// TIA Portal V20 export
// export: Created 2026-10-11T05:25:30.6576364Z, ExportSetting WithDefaults, DisplayName Totally Integrated Automation Portal, DisplayVersion V20, DisplayName TIA Portal Openness, DisplayVersion V20, DisplayName TIA Portal Teamcenter Gateway, DisplayVersion V20, DisplayName TIA Portal Version Control Interface, DisplayVersion V20, DisplayName SINAMICS Startdrive Advanced, DisplayVersion V20 SP1 Update 2, DisplayName SINAMICS Startdrive G110M, G120, G120C, G120D, G120P, G115D, DisplayVersion V20 SP1 Update 2, DisplayName SINAMICS Startdrive G130, G150, S120, S150, SINAMICS MV, G220, S200, S210, DisplayVersion V20 SP1 Update 2, DisplayName STEP 7 Professional, DisplayVersion V20, DisplayName STEP 7 Safety, DisplayVersion V20, DisplayName WinCC Basic/Comfort/Advanced, DisplayVersion V20, DisplayName WinCC Professional, DisplayVersion V20, DisplayName WinCC Unified, DisplayVersion V20
FUNCTION "FRK_PartReceived" : Bool   // FC38, SCL
{ S7_Optimized_Access := 'TRUE' }
VERSION : 0.1
// stored: AutoNumber true, IsIECCheckEnabled false, SetENOAutomatically false, UDAEnableTagReadback false
   VAR_IN_OUT
      Core : "FRK_Core";
      Unit : "FRK_Unit";
      Status : "ST_ModuleStatus";
      Part : "ST_PartContext";
      History : Array[1..16] of "ST_Diagnostic";
      Head : Int;
   END_VAR
   VAR_TEMP
      Index : DInt;
      Uid : String[64];
      ResultIndex : DInt;
   END_VAR
BEGIN

   #FRK_PartReceived := FALSE;
   #Index := #Unit.CarrierIndex;
   IF #Index = 0 THEN
       RETURN;
   END_IF;
   IF #Index < 1 OR #Index > 32 THEN
       "FRK_Fault"(Core := #Core,
                   Status := #Status,
                   ReasonCode := 2020,
                   Description := WSTRING#'std.error.partCarrierReadFailed');
       RETURN;
   END_IF;
   IF NOT "FRK_Carriers".Slots[#Index].Enabled OR "FRK_Carriers".Slots[#Index].Kind <> 2 OR "FRK_Carriers".Slots[#Index].Serial = UDINT#4294967295 THEN
       "FRK_Fault"(Core := #Core,
                   Status := #Status,
                   ReasonCode := 2020,
                   Description := WSTRING#'std.error.partCarrierReadFailed');
       RETURN;
   END_IF;
   "FRK_Carriers".Slots[#Index].Serial := "FRK_Carriers".Slots[#Index].Serial + 1;
   #Uid := CONCAT(IN1 := 'FRK-', IN2 := DINT_TO_STRING(#Index));
   #Uid := CONCAT(IN1 := #Uid, IN2 := '-');
   #Uid := CONCAT(IN1 := #Uid, IN2 := UDINT_TO_STRING("FRK_Carriers".Slots[#Index].Serial));
   #Part.Uid := #Uid;
   #Part.Present := TRUE;
   #Part.CarrierKind := 2;
   #Part.Result.Verdict := 0;
   #Part.Result.ReasonCode := 0;
   #Part.Result.StationPath := STRING_TO_WSTRING(#Status.Name);
   #Part.Result.Stamp := LDT#1970-01-01-00:00:00.000000000;
   #Part.Result.TimeSynchronized := FALSE;
   FOR #ResultIndex := 1 TO 32 DO
       #Part.Result.Records[#ResultIndex].Name := '';
   END_FOR;
   FOR #ResultIndex := 1 TO 8 DO
       #Part.Parents[#ResultIndex] := '';
   END_FOR;
   "FRK_Carriers".Slots[#Index].Context := #Part;
   "FRK_PartEvent"(History := #History,
                   Head := #Head,
                   Reason := 2024,
                   Uid := #Part.Uid,
                   SourcePath := #Status.Name);
   #FRK_PartReceived := TRUE;
END_FUNCTION
